DATA_BLOCK "ControlNodes"
{ S7_Optimized_Access := 'TRUE' }
VERSION : 0.1
NON_RETAIN
STRUCT
    sequence : "LAF_typeSequence";
    jobs : "LAF_typeJobs";
    cylFC2600FTControlFeed : "LBC_TwoWayActuatorControlNodes";
    sensorFC2600FTControlReady : "LBC_DigitalSignalControlNodes";
END_STRUCT;
BEGIN
END_DATA_BLOCK
